(* IEC 61131-3 sources: Versio-VersionControlSystem/fixtures/projects/RefrigeratorControl/Device/Plc Logic/Application/Library/Alarm/POUs/FB_Alarm/Private, 4 files *)

(* ---- _M_StateMachine.st ---- *)
METHOD PRIVATE _M_StateMachine

// --- BEGIN IMPLEMENTATION ---

// Alarm disabled
IF NOT Settings.Enable OR (NOT Condition AND State = E_AlarmState.Off) THEN
	RETURN;
END_IF

// State Machine
CASE State OF
	E_AlarmState.Off:
		IF DelayTimer.Q THEN
			NextState := E_AlarmState.Active;
		END_IF
	E_AlarmState.Active:
		IF DelayTimer.Q THEN
			NextState := E_AlarmState.Off;
		END_IF
	ELSE
		NextState := E_AlarmState.Off;
END_CASE

// Update State
_M_UpdateState();

(* ---- _M_UpdateState.st ---- *)
METHOD PRIVATE _M_UpdateState : BOOL

// --- BEGIN IMPLEMENTATION ---

// Update State
IF NextState <> State THEN
	State := NextState;

	//ResetTimer
	DelayTimer(IN := FALSE);

	IF State = E_AlarmState.Off THEN
		;//Configuration.Info := '';
	END_IF
END_IF

(* ---- _M_UpdateStatus.st ---- *)
METHOD PRIVATE _M_UpdateStatus : BOOL
VAR_INPUT
END_VAR

// --- BEGIN IMPLEMENTATION ---

(* ---- _M_EvaluateInputs.st ---- *)
METHOD PRIVATE _M_EvaluateInputs : BOOL
VAR_INST
	EnableRTrig	: R_TRIG;
	EnableFTrig	: F_TRIG;
END_VAR

// --- BEGIN IMPLEMENTATION ---

// Initialized
IF Settings.ShortDesc <> '' AND NOT Configuration.Initialized THEN
	Configuration.Initialized := TRUE;
END_IF

// Enable State change
EnableRTrig(CLK := Settings.Enable);
EnableFTrig(CLK := Settings.Enable);
IF EnableRTrig.Q OR EnableFTrig.Q THEN
	NextState := E_AlarmState.Off;
	_M_UpdateState();
END_IF

// Delays
_M_Timers();
